// --- Siemens Structured Format ---
DATA_BLOCK "model__HS8_IW100_"
{ S7_Optimized_Access := 'TRUE' }
VERSION :
NON_RETAIN
   VAR
      W_i : ARRAY[0..7, 0..39] OF REAL;
      W_f : ARRAY[0..7, 0..39] OF REAL;
      W_g : ARRAY[0..7, 0..39] OF REAL;
      W_o : ARRAY[0..7, 0..39] OF REAL;
      R_i : ARRAY[0..7, 0..7] OF REAL;
      R_f : ARRAY[0..7, 0..7] OF REAL;
      R_g : ARRAY[0..7, 0..7] OF REAL;
      R_o : ARRAY[0..7, 0..7] OF REAL;
      B_i : ARRAY[0..7] OF REAL;
      B_f : ARRAY[0..7] OF REAL;
      B_g : ARRAY[0..7] OF REAL;
      B_o : ARRAY[0..7] OF REAL;
      FC_W : ARRAY[0..39, 0..7] OF REAL;
      FC_B : ARRAY[0..39] OF REAL;
   END_VAR
BEGIN

      W_i[0,0] := -0.00829199;
      W_i[0,1] := 0.04314763;
      W_i[0,2] := -0.00093121;
      W_i[0,3] := -0.41203406;
      W_i[0,4] := 0.14360030;
      W_i[0,5] := -0.00333697;
      W_i[0,6] := -0.05594388;
      W_i[0,7] := 0.22901678;
      W_i[0,8] := 0.12452386;
      W_i[0,9] := 0.18269505;
      W_i[0,10] := -0.00489003;
      W_i[0,11] := -1.12929618;
      W_i[0,12] := 0.50561267;
      W_i[0,13] := -0.01176495;
      W_i[0,14] := 0.05196610;
      W_i[0,15] := 0.29604533;
      W_i[0,16] := 0.00854590;
      W_i[0,17] := 0.00023653;
      W_i[0,18] := -0.05930486;
      W_i[0,19] := 0.34416831;
      W_i[0,20] := 0.04249638;
      W_i[0,21] := 0.29057521;
      W_i[0,22] := 0.00544647;
      W_i[0,23] := -0.19255431;
      W_i[0,24] := -0.20954449;
      W_i[0,25] := -0.09120649;
      W_i[0,26] := -0.00158587;
      W_i[0,27] := -0.21091045;
      W_i[0,28] := -0.00354010;
      W_i[0,29] := -0.11485449;
      W_i[0,30] := 0.40112287;
      W_i[0,31] := -0.23464951;
      W_i[0,32] := 0.07507721;
      W_i[0,33] := -0.04070815;
      W_i[0,34] := 0.16331266;
      W_i[0,35] := -0.06922071;
      W_i[0,36] := 0.07785974;
      W_i[0,37] := -0.12469714;
      W_i[0,38] := -0.09480914;
      W_i[0,39] := -0.12007505;
      W_i[1,0] := -0.14511052;
      W_i[1,1] := 0.01258339;
      W_i[1,2] := -0.02499544;
      W_i[1,3] := -0.02792050;
      W_i[1,4] := 0.05153107;
      W_i[1,5] := 0.02871069;
      W_i[1,6] := -0.00801326;
      W_i[1,7] := 0.16971111;
      W_i[1,8] := 0.07463019;
      W_i[1,9] := -0.30484986;
      W_i[1,10] := 0.00891454;
      W_i[1,11] := 0.19871780;
      W_i[1,12] := 0.02821600;
      W_i[1,13] := -0.07369927;
      W_i[1,14] := 0.02203551;
      W_i[1,15] := 0.08398883;
      W_i[1,16] := 0.00458911;
      W_i[1,17] := 0.01521466;
      W_i[1,18] := 0.06061148;
      W_i[1,19] := -0.08532640;
      W_i[1,20] := 0.01589951;
      W_i[1,21] := 0.00234504;
      W_i[1,22] := -0.04496472;
      W_i[1,23] := -0.04576229;
      W_i[1,24] := 0.03349697;
      W_i[1,25] := -0.14834076;
      W_i[1,26] := -0.00671506;
      W_i[1,27] := -0.04002256;
      W_i[1,28] := -0.05524301;
      W_i[1,29] := -0.04596998;
      W_i[1,30] := 0.20154108;
      W_i[1,31] := -0.04227936;
      W_i[1,32] := 0.27783859;
      W_i[1,33] := -0.15889524;
      W_i[1,34] := -0.17870863;
      W_i[1,35] := -0.22829576;
      W_i[1,36] := 0.00769149;
      W_i[1,37] := 0.21033208;
      W_i[1,38] := 0.02056267;
      W_i[1,39] := 0.03890164;
      W_i[2,0] := -0.00940658;
      W_i[2,1] := 0.01171005;
      W_i[2,2] := 0.01976776;
      W_i[2,3] := -0.01506334;
      W_i[2,4] := -0.01478560;
      W_i[2,5] := 0.02109193;
      W_i[2,6] := 0.01444429;
      W_i[2,7] := 0.00977760;
      W_i[2,8] := 0.06673528;
      W_i[2,9] := 0.07852798;
      W_i[2,10] := -0.02388507;
      W_i[2,11] := 0.15636960;
      W_i[2,12] := 0.04547270;
      W_i[2,13] := 0.05332979;
      W_i[2,14] := 0.02128568;
      W_i[2,15] := -0.06670643;
      W_i[2,16] := -0.00303149;
      W_i[2,17] := -0.01812665;
      W_i[2,18] := 0.09366660;
      W_i[2,19] := -0.02572775;
      W_i[2,20] := -0.02855127;
      W_i[2,21] := -0.05881069;
      W_i[2,22] := -0.05029222;
      W_i[2,23] := 0.09357284;
      W_i[2,24] := -0.46770903;
      W_i[2,25] := -0.71739095;
      W_i[2,26] := -0.03358178;
      W_i[2,27] := -0.11196791;
      W_i[2,28] := 0.12867627;
      W_i[2,29] := -0.15594745;
      W_i[2,30] := -0.02176742;
      W_i[2,31] := 0.05814255;
      W_i[2,32] := 0.02967955;
      W_i[2,33] := -0.32135192;
      W_i[2,34] := -0.70631939;
      W_i[2,35] := 0.13404904;
      W_i[2,36] := -0.05614626;
      W_i[2,37] := -0.06990065;
      W_i[2,38] := 0.09054608;
      W_i[2,39] := 0.08889610;
      W_i[3,0] := 0.05596327;
      W_i[3,1] := -0.32603350;
      W_i[3,2] := -0.13964993;
      W_i[3,3] := -0.15204740;
      W_i[3,4] := 0.05851153;
      W_i[3,5] := 0.08759125;
      W_i[3,6] := 0.07076695;
      W_i[3,7] := 0.05082684;
      W_i[3,8] := 0.00611771;
      W_i[3,9] := -0.05680722;
      W_i[3,10] := 0.04656018;
      W_i[3,11] := 0.08742622;
      W_i[3,12] := -0.00764282;
      W_i[3,13] := -0.35034382;
      W_i[3,14] := -0.12616983;
      W_i[3,15] := 0.03790347;
      W_i[3,16] := -0.00427554;
      W_i[3,17] := 0.10194600;
      W_i[3,18] := -0.06467836;
      W_i[3,19] := -0.04557304;
      W_i[3,20] := 0.13014187;
      W_i[3,21] := -0.11706656;
      W_i[3,22] := 0.20328589;
      W_i[3,23] := 0.31214345;
      W_i[3,24] := -0.19055620;
      W_i[3,25] := 0.11225392;
      W_i[3,26] := -0.00316885;
      W_i[3,27] := 0.02801218;
      W_i[3,28] := 0.07838947;
      W_i[3,29] := -0.08224142;
      W_i[3,30] := 0.02575504;
      W_i[3,31] := 0.07745822;
      W_i[3,32] := 0.05140261;
      W_i[3,33] := 0.00126193;
      W_i[3,34] := 0.03769523;
      W_i[3,35] := -0.21655150;
      W_i[3,36] := -0.08745287;
      W_i[3,37] := 0.10195030;
      W_i[3,38] := -0.44626316;
      W_i[3,39] := -0.86872011;
      W_i[4,0] := -0.04617658;
      W_i[4,1] := -0.03314103;
      W_i[4,2] := -0.08659177;
      W_i[4,3] := -0.10351395;
      W_i[4,4] := 0.06772576;
      W_i[4,5] := -0.04269263;
      W_i[4,6] := -0.04438864;
      W_i[4,7] := -0.01167864;
      W_i[4,8] := 0.02057231;
      W_i[4,9] := -0.07837452;
      W_i[4,10] := -0.03820154;
      W_i[4,11] := -0.03692231;
      W_i[4,12] := -0.07637376;
      W_i[4,13] := -0.06241865;
      W_i[4,14] := -0.01509702;
      W_i[4,15] := 0.07582836;
      W_i[4,16] := -0.01766248;
      W_i[4,17] := 0.00024068;
      W_i[4,18] := 0.03632537;
      W_i[4,19] := 0.01485146;
      W_i[4,20] := 0.10803255;
      W_i[4,21] := -0.14425407;
      W_i[4,22] := -0.01218021;
      W_i[4,23] := -0.01190184;
      W_i[4,24] := -0.46979687;
      W_i[4,25] := -0.46851084;
      W_i[4,26] := -0.02849982;
      W_i[4,27] := 0.03427306;
      W_i[4,28] := 0.04523883;
      W_i[4,29] := 0.25723371;
      W_i[4,30] := -0.09724599;
      W_i[4,31] := 0.03623974;
      W_i[4,32] := -0.10095317;
      W_i[4,33] := 0.12443283;
      W_i[4,34] := -0.42049277;
      W_i[4,35] := -0.03480925;
      W_i[4,36] := 0.04771702;
      W_i[4,37] := 0.04326405;
      W_i[4,38] := 0.03356932;
      W_i[4,39] := 0.03849664;
      W_i[5,0] := -0.17091992;
      W_i[5,1] := -0.04787771;
      W_i[5,2] := -0.02202379;
      W_i[5,3] := -0.09034166;
      W_i[5,4] := -0.00740036;
      W_i[5,5] := 0.00184778;
      W_i[5,6] := 0.01398086;
      W_i[5,7] := -0.08714975;
      W_i[5,8] := -0.10723638;
      W_i[5,9] := 0.27444202;
      W_i[5,10] := 0.02795951;
      W_i[5,11] := 0.16468486;
      W_i[5,12] := -0.25734791;
      W_i[5,13] := -0.08599530;
      W_i[5,14] := -0.07228005;
      W_i[5,15] := 0.24830806;
      W_i[5,16] := 0.04241711;
      W_i[5,17] := -0.00679267;
      W_i[5,18] := 1.35323977;
      W_i[5,19] := 0.07199069;
      W_i[5,20] := 0.06845883;
      W_i[5,21] := 0.20864677;
      W_i[5,22] := -0.14911477;
      W_i[5,23] := 0.14023533;
      W_i[5,24] := -0.02367306;
      W_i[5,25] := 0.60291624;
      W_i[5,26] := -0.19428003;
      W_i[5,27] := -0.32415670;
      W_i[5,28] := 0.17960674;
      W_i[5,29] := 0.09058087;
      W_i[5,30] := -0.24361624;
      W_i[5,31] := -0.07183243;
      W_i[5,32] := 0.01278071;
      W_i[5,33] := -0.11311200;
      W_i[5,34] := 0.64622027;
      W_i[5,35] := -0.06918935;
      W_i[5,36] := 0.04555825;
      W_i[5,37] := -0.41487035;
      W_i[5,38] := -0.02093678;
      W_i[5,39] := 0.11062510;
      W_i[6,0] := -0.08444463;
      W_i[6,1] := 0.03796263;
      W_i[6,2] := 0.02793699;
      W_i[6,3] := 0.08258326;
      W_i[6,4] := 0.01806726;
      W_i[6,5] := 0.04154406;
      W_i[6,6] := 0.06518649;
      W_i[6,7] := -0.35571000;
      W_i[6,8] := -0.08575057;
      W_i[6,9] := 0.03024576;
      W_i[6,10] := 0.08267769;
      W_i[6,11] := -0.51406556;
      W_i[6,12] := -0.18283555;
      W_i[6,13] := 0.08692829;
      W_i[6,14] := -0.01571506;
      W_i[6,15] := 0.41990465;
      W_i[6,16] := 0.06421173;
      W_i[6,17] := 0.02368255;
      W_i[6,18] := 0.00736057;
      W_i[6,19] := 0.13490863;
      W_i[6,20] := 0.24439722;
      W_i[6,21] := 0.22145407;
      W_i[6,22] := 0.23587099;
      W_i[6,23] := -0.08479463;
      W_i[6,24] := 0.15434107;
      W_i[6,25] := 0.35517022;
      W_i[6,26] := 0.02139992;
      W_i[6,27] := -0.18648548;
      W_i[6,28] := 0.00971483;
      W_i[6,29] := -0.15883411;
      W_i[6,30] := 0.16745885;
      W_i[6,31] := -0.09647866;
      W_i[6,32] := 0.20241226;
      W_i[6,33] := -0.10213183;
      W_i[6,34] := 0.35625863;
      W_i[6,35] := -0.21271712;
      W_i[6,36] := 0.07117779;
      W_i[6,37] := -0.05264070;
      W_i[6,38] := -0.07197802;
      W_i[6,39] := 0.05570221;
      W_i[7,0] := -0.14402835;
      W_i[7,1] := -0.07068059;
      W_i[7,2] := 0.04391022;
      W_i[7,3] := -0.23145308;
      W_i[7,4] := 0.01739045;
      W_i[7,5] := -0.09847571;
      W_i[7,6] := -0.07244503;
      W_i[7,7] := 0.54241705;
      W_i[7,8] := 0.05786600;
      W_i[7,9] := -0.11313851;
      W_i[7,10] := 0.05011918;
      W_i[7,11] := -0.88967866;
      W_i[7,12] := -0.78758240;
      W_i[7,13] := -0.07027908;
      W_i[7,14] := -0.15626858;
      W_i[7,15] := -0.01163841;
      W_i[7,16] := 0.06607775;
      W_i[7,17] := -0.20021817;
      W_i[7,18] := 0.08560139;
      W_i[7,19] := -0.06735905;
      W_i[7,20] := 0.11073713;
      W_i[7,21] := 0.03392316;
      W_i[7,22] := -0.07517586;
      W_i[7,23] := -0.07473031;
      W_i[7,24] := 0.17482267;
      W_i[7,25] := 0.75477821;
      W_i[7,26] := -0.19560531;
      W_i[7,27] := -0.00529976;
      W_i[7,28] := 0.06779508;
      W_i[7,29] := -0.05984003;
      W_i[7,30] := 0.36871162;
      W_i[7,31] := 0.09751310;
      W_i[7,32] := -0.32882604;
      W_i[7,33] := 0.10271895;
      W_i[7,34] := 0.03595359;
      W_i[7,35] := -0.06912012;
      W_i[7,36] := 0.05955562;
      W_i[7,37] := 0.15649518;
      W_i[7,38] := -0.16574396;
      W_i[7,39] := 0.02650662;
      W_f[0,0] := -0.08104721;
      W_f[0,1] := 0.02299085;
      W_f[0,2] := -0.08156814;
      W_f[0,3] := 0.34981409;
      W_f[0,4] := -0.02991411;
      W_f[0,5] := 0.05847026;
      W_f[0,6] := 0.08058469;
      W_f[0,7] := 0.08683547;
      W_f[0,8] := 0.02113942;
      W_f[0,9] := -0.22806560;
      W_f[0,10] := -0.04616724;
      W_f[0,11] := -0.04299140;
      W_f[0,12] := 0.11675275;
      W_f[0,13] := -0.09660369;
      W_f[0,14] := -0.04888760;
      W_f[0,15] := -0.18213840;
      W_f[0,16] := 0.12695764;
      W_f[0,17] := 0.22833031;
      W_f[0,18] := -0.03068344;
      W_f[0,19] := -0.22004378;
      W_f[0,20] := 0.01699636;
      W_f[0,21] := 0.10058182;
      W_f[0,22] := 0.02436358;
      W_f[0,23] := 0.01155086;
      W_f[0,24] := 0.67554194;
      W_f[0,25] := 0.77170414;
      W_f[0,26] := 0.04872859;
      W_f[0,27] := 0.04316394;
      W_f[0,28] := 0.01004832;
      W_f[0,29] := 0.10533538;
      W_f[0,30] := 0.26388049;
      W_f[0,31] := 0.16926253;
      W_f[0,32] := 0.31521299;
      W_f[0,33] := 0.23292090;
      W_f[0,34] := 0.71050066;
      W_f[0,35] := 0.07673426;
      W_f[0,36] := -0.03209021;
      W_f[0,37] := -0.07602870;
      W_f[0,38] := 0.07363247;
      W_f[0,39] := 0.09119339;
      W_f[1,0] := -0.02197713;
      W_f[1,1] := -0.01616614;
      W_f[1,2] := -0.02013298;
      W_f[1,3] := -0.00875140;
      W_f[1,4] := 0.04112979;
      W_f[1,5] := 0.05162001;
      W_f[1,6] := 0.00973919;
      W_f[1,7] := 0.07910040;
      W_f[1,8] := -0.31076026;
      W_f[1,9] := 0.18630370;
      W_f[1,10] := -0.00576194;
      W_f[1,11] := 0.04994554;
      W_f[1,12] := 0.05406393;
      W_f[1,13] := 0.05481998;
      W_f[1,14] := 0.01417492;
      W_f[1,15] := -0.11486354;
      W_f[1,16] := 0.22028089;
      W_f[1,17] := 0.03549247;
      W_f[1,18] := 0.07496776;
      W_f[1,19] := -0.31716284;
      W_f[1,20] := 0.02977121;
      W_f[1,21] := -0.10077871;
      W_f[1,22] := 0.29007021;
      W_f[1,23] := 0.02756922;
      W_f[1,24] := 1.14809716;
      W_f[1,25] := 1.46478581;
      W_f[1,26] := -0.01241822;
      W_f[1,27] := 0.09172244;
      W_f[1,28] := 0.01175412;
      W_f[1,29] := -0.10488217;
      W_f[1,30] := 0.00364918;
      W_f[1,31] := -0.03901139;
      W_f[1,32] := -0.08511472;
      W_f[1,33] := 0.08891900;
      W_f[1,34] := 1.39858294;
      W_f[1,35] := -0.42813861;
      W_f[1,36] := -0.00882304;
      W_f[1,37] := -0.05784527;
      W_f[1,38] := -0.13634762;
      W_f[1,39] := 0.17077002;
      W_f[2,0] := 0.01542370;
      W_f[2,1] := 0.01987428;
      W_f[2,2] := 0.00323933;
      W_f[2,3] := -0.01730455;
      W_f[2,4] := 0.06355638;
      W_f[2,5] := 0.03613569;
      W_f[2,6] := -0.01693674;
      W_f[2,7] := -0.01970888;
      W_f[2,8] := -0.06606199;
      W_f[2,9] := -0.07453630;
      W_f[2,10] := -0.00336948;
      W_f[2,11] := -0.20352897;
      W_f[2,12] := -0.10294267;
      W_f[2,13] := 0.02081121;
      W_f[2,14] := 0.06329557;
      W_f[2,15] := 0.02846926;
      W_f[2,16] := 0.06616816;
      W_f[2,17] := 0.00726432;
      W_f[2,18] := 0.04505518;
      W_f[2,19] := 0.02842713;
      W_f[2,20] := -0.00391449;
      W_f[2,21] := -0.00121696;
      W_f[2,22] := -0.17400308;
      W_f[2,23] := 0.02276708;
      W_f[2,24] := 0.26592869;
      W_f[2,25] := 0.03894256;
      W_f[2,26] := 0.12431550;
      W_f[2,27] := -0.02150069;
      W_f[2,28] := -0.05582710;
      W_f[2,29] := 0.25016540;
      W_f[2,30] := 0.01012970;
      W_f[2,31] := -0.01360032;
      W_f[2,32] := -0.07151139;
      W_f[2,33] := 0.20726912;
      W_f[2,34] := -0.33328736;
      W_f[2,35] := 0.15157171;
      W_f[2,36] := 0.01685908;
      W_f[2,37] := -0.12045209;
      W_f[2,38] := 0.01227041;
      W_f[2,39] := 0.06517339;
      W_f[3,0] := 0.47573653;
      W_f[3,1] := 0.13755870;
      W_f[3,2] := -0.08410271;
      W_f[3,3] := -0.16147336;
      W_f[3,4] := 0.10956663;
      W_f[3,5] := -0.05382008;
      W_f[3,6] := -0.09864125;
      W_f[3,7] := 0.37438312;
      W_f[3,8] := -0.31137553;
      W_f[3,9] := 0.11690006;
      W_f[3,10] := -0.16711678;
      W_f[3,11] := -0.35226113;
      W_f[3,12] := 0.14284903;
      W_f[3,13] := 0.22532572;
      W_f[3,14] := 0.31750289;
      W_f[3,15] := -0.04833202;
      W_f[3,16] := 0.04104101;
      W_f[3,17] := -0.29455543;
      W_f[3,18] := -2.66076255;
      W_f[3,19] := -0.09576055;
      W_f[3,20] := -0.16356435;
      W_f[3,21] := 0.10903085;
      W_f[3,22] := -0.44664004;
      W_f[3,23] := -0.17856193;
      W_f[3,24] := 0.41079015;
      W_f[3,25] := 0.15273106;
      W_f[3,26] := -0.33044237;
      W_f[3,27] := -0.18228154;
      W_f[3,28] := 0.04568926;
      W_f[3,29] := 1.02778792;
      W_f[3,30] := -0.34178400;
      W_f[3,31] := -0.00056406;
      W_f[3,32] := 0.21154980;
      W_f[3,33] := -0.10385001;
      W_f[3,34] := 0.03440418;
      W_f[3,35] := 0.25746328;
      W_f[3,36] := 0.02392143;
      W_f[3,37] := -0.14384723;
      W_f[3,38] := 0.40537423;
      W_f[3,39] := -0.08356514;
      W_f[4,0] := 0.01179661;
      W_f[4,1] := 0.06130485;
      W_f[4,2] := 0.00775665;
      W_f[4,3] := -0.01987305;
      W_f[4,4] := 0.03156713;
      W_f[4,5] := -0.03151586;
      W_f[4,6] := -0.06941684;
      W_f[4,7] := -0.05865467;
      W_f[4,8] := -0.12223195;
      W_f[4,9] := 0.00069460;
      W_f[4,10] := -0.01235222;
      W_f[4,11] := -0.05694751;
      W_f[4,12] := -0.00690056;
      W_f[4,13] := 0.02081548;
      W_f[4,14] := -0.02345082;
      W_f[4,15] := -0.08427138;
      W_f[4,16] := 0.00219320;
      W_f[4,17] := -0.00790089;
      W_f[4,18] := 0.06579314;
      W_f[4,19] := -0.04613130;
      W_f[4,20] := 0.06156648;
      W_f[4,21] := 0.08230194;
      W_f[4,22] := 0.02192603;
      W_f[4,23] := -0.05004644;
      W_f[4,24] := -0.33776584;
      W_f[4,25] := -0.57119745;
      W_f[4,26] := 0.00284863;
      W_f[4,27] := -0.03237003;
      W_f[4,28] := -0.06698364;
      W_f[4,29] := -0.32339925;
      W_f[4,30] := 0.06599762;
      W_f[4,31] := 0.03372506;
      W_f[4,32] := 0.20183899;
      W_f[4,33] := 0.09781818;
      W_f[4,34] := 0.21647416;
      W_f[4,35] := -0.03968338;
      W_f[4,36] := 0.04764435;
      W_f[4,37] := -0.09999206;
      W_f[4,38] := -0.04979988;
      W_f[4,39] := 0.04298165;
      W_f[5,0] := -0.00328023;
      W_f[5,1] := 0.05526555;
      W_f[5,2] := -0.02378737;
      W_f[5,3] := 0.07470135;
      W_f[5,4] := 0.07415909;
      W_f[5,5] := 0.03875844;
      W_f[5,6] := 0.04064441;
      W_f[5,7] := 0.01137258;
      W_f[5,8] := 0.04157886;
      W_f[5,9] := -0.11250745;
      W_f[5,10] := -0.03683221;
      W_f[5,11] := -0.05140235;
      W_f[5,12] := 0.16510846;
      W_f[5,13] := -0.00409127;
      W_f[5,14] := -0.03037189;
      W_f[5,15] := -0.14330336;
      W_f[5,16] := -0.02087791;
      W_f[5,17] := 0.05005715;
      W_f[5,18] := -0.06411071;
      W_f[5,19] := -0.05833034;
      W_f[5,20] := 0.00247585;
      W_f[5,21] := 0.07365038;
      W_f[5,22] := 0.00771155;
      W_f[5,23] := -0.07253324;
      W_f[5,24] := 0.94747639;
      W_f[5,25] := 0.65536422;
      W_f[5,26] := 0.01926010;
      W_f[5,27] := -0.07741715;
      W_f[5,28] := -0.02838454;
      W_f[5,29] := -0.25596547;
      W_f[5,30] := 0.04823640;
      W_f[5,31] := 0.03441899;
      W_f[5,32] := -0.04197009;
      W_f[5,33] := 0.14078745;
      W_f[5,34] := 0.25478148;
      W_f[5,35] := -0.08758619;
      W_f[5,36] := -0.00409188;
      W_f[5,37] := 0.10015804;
      W_f[5,38] := -0.01840312;
      W_f[5,39] := 0.04281899;
      W_f[6,0] := -0.03747290;
      W_f[6,1] := 0.00117479;
      W_f[6,2] := 0.01929842;
      W_f[6,3] := -0.16080324;
      W_f[6,4] := -0.00967213;
      W_f[6,5] := 0.02158868;
      W_f[6,6] := -0.07005120;
      W_f[6,7] := 0.21899310;
      W_f[6,8] := 0.03782399;
      W_f[6,9] := -0.21971041;
      W_f[6,10] := -0.04937140;
      W_f[6,11] := 0.04276552;
      W_f[6,12] := 0.02347153;
      W_f[6,13] := -0.08741955;
      W_f[6,14] := 0.02819359;
      W_f[6,15] := -0.32513508;
      W_f[6,16] := 0.09819235;
      W_f[6,17] := -0.00175993;
      W_f[6,18] := 0.00046430;
      W_f[6,19] := 0.00414359;
      W_f[6,20] := 0.05726501;
      W_f[6,21] := 0.02174316;
      W_f[6,22] := 0.40702432;
      W_f[6,23] := 0.05224282;
      W_f[6,24] := 1.36585915;
      W_f[6,25] := 1.40137434;
      W_f[6,26] := 0.06176697;
      W_f[6,27] := 0.03423437;
      W_f[6,28] := 0.01783603;
      W_f[6,29] := -0.56917655;
      W_f[6,30] := 0.47907564;
      W_f[6,31] := 0.10644426;
      W_f[6,32] := 0.44268256;
      W_f[6,33] := 0.56317347;
      W_f[6,34] := 1.12857997;
      W_f[6,35] := 0.00323946;
      W_f[6,36] := -0.03574727;
      W_f[6,37] := -0.12019916;
      W_f[6,38] := -0.04353496;
      W_f[6,39] := 0.18841393;
      W_f[7,0] := 0.08367904;
      W_f[7,1] := -0.02769166;
      W_f[7,2] := 0.05256313;
      W_f[7,3] := -0.02467708;
      W_f[7,4] := -0.08298105;
      W_f[7,5] := -0.01648388;
      W_f[7,6] := -0.04057755;
      W_f[7,7] := 0.05192674;
      W_f[7,8] := -0.03598220;
      W_f[7,9] := -0.13019682;
      W_f[7,10] := 0.01959694;
      W_f[7,11] := 0.00413586;
      W_f[7,12] := 0.05873092;
      W_f[7,13] := 0.02881050;
      W_f[7,14] := -0.02888235;
      W_f[7,15] := -0.13839944;
      W_f[7,16] := 0.02485734;
      W_f[7,17] := -0.11965133;
      W_f[7,18] := -0.11112632;
      W_f[7,19] := 0.03353542;
      W_f[7,20] := 0.02333037;
      W_f[7,21] := 0.04703392;
      W_f[7,22] := 0.20441540;
      W_f[7,23] := 0.07088239;
      W_f[7,24] := 0.59273797;
      W_f[7,25] := 0.38002837;
      W_f[7,26] := 0.01679641;
      W_f[7,27] := 0.03724186;
      W_f[7,28] := -0.06413292;
      W_f[7,29] := -0.13961390;
      W_f[7,30] := 0.11306310;
      W_f[7,31] := -0.00102062;
      W_f[7,32] := 0.19089061;
      W_f[7,33] := 0.12474129;
      W_f[7,34] := 0.52092993;
      W_f[7,35] := 0.02751438;
      W_f[7,36] := 0.01992416;
      W_f[7,37] := -0.08247742;
      W_f[7,38] := -0.05664129;
      W_f[7,39] := 0.16597328;
      W_g[0,0] := -0.06630491;
      W_g[0,1] := 0.02753393;
      W_g[0,2] := -0.06609154;
      W_g[0,3] := 0.03565337;
      W_g[0,4] := -0.14254735;
      W_g[0,5] := 0.07333323;
      W_g[0,6] := 0.14428975;
      W_g[0,7] := 0.03311217;
      W_g[0,8] := 0.02892466;
      W_g[0,9] := 0.04255950;
      W_g[0,10] := -0.03547552;
      W_g[0,11] := 0.02729788;
      W_g[0,12] := 0.02407304;
      W_g[0,13] := -0.01838484;
      W_g[0,14] := -0.04254790;
      W_g[0,15] := 0.00052823;
      W_g[0,16] := 0.02627059;
      W_g[0,17] := 0.12881427;
      W_g[0,18] := -0.04993503;
      W_g[0,19] := 0.05080932;
      W_g[0,20] := -0.13986340;
      W_g[0,21] := 0.11638415;
      W_g[0,22] := 0.01129120;
      W_g[0,23] := -0.00916141;
      W_g[0,24] := 0.20254859;
      W_g[0,25] := 0.08704451;
      W_g[0,26] := -0.03924693;
      W_g[0,27] := 0.10738914;
      W_g[0,28] := -0.04623365;
      W_g[0,29] := -0.00351558;
      W_g[0,30] := 0.00354978;
      W_g[0,31] := 0.00794905;
      W_g[0,32] := 0.00442744;
      W_g[0,33] := 0.00612418;
      W_g[0,34] := -0.20538065;
      W_g[0,35] := 0.03906323;
      W_g[0,36] := -0.00062364;
      W_g[0,37] := 0.00209236;
      W_g[0,38] := -0.03761620;
      W_g[0,39] := -0.04062740;
      W_g[1,0] := -0.10235135;
      W_g[1,1] := 0.06025442;
      W_g[1,2] := -0.09398326;
      W_g[1,3] := 0.05591756;
      W_g[1,4] := -0.10170189;
      W_g[1,5] := 0.04167721;
      W_g[1,6] := 0.01649847;
      W_g[1,7] := 0.04434075;
      W_g[1,8] := 0.04717555;
      W_g[1,9] := 0.03831566;
      W_g[1,10] := 0.05404275;
      W_g[1,11] := 0.16338016;
      W_g[1,12] := 0.15951122;
      W_g[1,13] := 0.02527176;
      W_g[1,14] := -0.01270708;
      W_g[1,15] := 0.16955729;
      W_g[1,16] := -0.08400796;
      W_g[1,17] := -0.09564576;
      W_g[1,18] := -0.16610350;
      W_g[1,19] := 0.18888752;
      W_g[1,20] := -0.02569673;
      W_g[1,21] := -0.05631816;
      W_g[1,22] := -0.01589629;
      W_g[1,23] := 0.06837284;
      W_g[1,24] := 0.19006948;
      W_g[1,25] := -0.18527375;
      W_g[1,26] := 0.06264018;
      W_g[1,27] := -0.06131431;
      W_g[1,28] := -0.02992554;
      W_g[1,29] := 0.02249875;
      W_g[1,30] := -0.01341370;
      W_g[1,31] := -0.01471063;
      W_g[1,32] := -0.01641031;
      W_g[1,33] := -0.02138708;
      W_g[1,34] := 0.09338091;
      W_g[1,35] := 0.17898178;
      W_g[1,36] := -0.08693415;
      W_g[1,37] := -0.19239108;
      W_g[1,38] := -0.05011347;
      W_g[1,39] := -0.03428216;
      W_g[2,0] := 0.06590919;
      W_g[2,1] := 0.01555668;
      W_g[2,2] := 0.05944061;
      W_g[2,3] := -0.00003379;
      W_g[2,4] := -0.16144016;
      W_g[2,5] := 0.07584924;
      W_g[2,6] := 0.07926709;
      W_g[2,7] := 0.00562621;
      W_g[2,8] := 0.00176247;
      W_g[2,9] := 0.00667630;
      W_g[2,10] := -0.01289325;
      W_g[2,11] := -0.03508691;
      W_g[2,12] := -0.03598065;
      W_g[2,13] := 0.14380608;
      W_g[2,14] := 0.06675316;
      W_g[2,15] := -0.02170967;
      W_g[2,16] := 0.03013330;
      W_g[2,17] := -0.04029799;
      W_g[2,18] := -0.14855465;
      W_g[2,19] := 0.00260400;
      W_g[2,20] := -0.08315958;
      W_g[2,21] := 0.01309617;
      W_g[2,22] := 0.05792306;
      W_g[2,23] := 0.14916992;
      W_g[2,24] := 0.13496941;
      W_g[2,25] := 0.20256528;
      W_g[2,26] := 0.06222376;
      W_g[2,27] := 0.00734210;
      W_g[2,28] := -0.04847896;
      W_g[2,29] := -0.00581570;
      W_g[2,30] := 0.03206468;
      W_g[2,31] := 0.02264830;
      W_g[2,32] := 0.04472146;
      W_g[2,33] := 0.04833479;
      W_g[2,34] := 0.68682790;
      W_g[2,35] := 0.03641244;
      W_g[2,36] := -0.05233013;
      W_g[2,37] := 0.01984018;
      W_g[2,38] := 0.05872162;
      W_g[2,39] := 0.05237507;
      W_g[3,0] := -0.05719843;
      W_g[3,1] := 0.06765803;
      W_g[3,2] := -0.05017579;
      W_g[3,3] := -0.09871275;
      W_g[3,4] := -0.14791933;
      W_g[3,5] := -0.05363221;
      W_g[3,6] := -0.11064304;
      W_g[3,7] := -0.06622731;
      W_g[3,8] := -0.06549069;
      W_g[3,9] := -0.07995880;
      W_g[3,10] := -0.00412930;
      W_g[3,11] := -0.05527864;
      W_g[3,12] := -0.05236278;
      W_g[3,13] := 0.01281861;
      W_g[3,14] := 0.00663725;
      W_g[3,15] := -0.05022956;
      W_g[3,16] := 0.00247445;
      W_g[3,17] := -0.00537014;
      W_g[3,18] := -0.17336990;
      W_g[3,19] := -0.04672612;
      W_g[3,20] := 0.08145336;
      W_g[3,21] := 0.04289828;
      W_g[3,22] := -0.04270948;
      W_g[3,23] := -0.00124830;
      W_g[3,24] := -0.58283401;
      W_g[3,25] := -0.74716926;
      W_g[3,26] := -0.05420419;
      W_g[3,27] := 0.04391639;
      W_g[3,28] := -0.21304598;
      W_g[3,29] := 0.14126062;
      W_g[3,30] := -0.04634099;
      W_g[3,31] := -0.01238058;
      W_g[3,32] := -0.02521331;
      W_g[3,33] := -0.01312026;
      W_g[3,34] := 0.00096928;
      W_g[3,35] := -0.08583874;
      W_g[3,36] := 0.04279795;
      W_g[3,37] := 0.07323888;
      W_g[3,38] := -0.00020507;
      W_g[3,39] := 0.48666921;
      W_g[4,0] := 0.03492008;
      W_g[4,1] := -0.06098935;
      W_g[4,2] := 0.03832612;
      W_g[4,3] := 0.05924186;
      W_g[4,4] := -0.04744076;
      W_g[4,5] := 0.03529921;
      W_g[4,6] := 0.07721187;
      W_g[4,7] := 0.05416005;
      W_g[4,8] := 0.05382877;
      W_g[4,9] := 0.06243544;
      W_g[4,10] := 0.00853686;
      W_g[4,11] := -0.00808500;
      W_g[4,12] := -0.00045702;
      W_g[4,13] := -0.01504347;
      W_g[4,14] := 0.05096063;
      W_g[4,15] := 0.00273409;
      W_g[4,16] := 0.04891136;
      W_g[4,17] := 0.01359798;
      W_g[4,18] := -0.04669548;
      W_g[4,19] := 0.01079443;
      W_g[4,20] := -0.08128674;
      W_g[4,21] := 0.02045462;
      W_g[4,22] := -0.03726062;
      W_g[4,23] := 0.01082981;
      W_g[4,24] := -0.72472757;
      W_g[4,25] := -0.60457122;
      W_g[4,26] := -0.02546896;
      W_g[4,27] := 0.02074758;
      W_g[4,28] := 0.02423066;
      W_g[4,29] := 0.02050022;
      W_g[4,30] := -0.03584260;
      W_g[4,31] := -0.03780675;
      W_g[4,32] := -0.01639182;
      W_g[4,33] := -0.01888406;
      W_g[4,34] := -0.90565455;
      W_g[4,35] := -0.02123658;
      W_g[4,36] := -0.05081832;
      W_g[4,37] := -0.08846542;
      W_g[4,38] := 0.05660410;
      W_g[4,39] := 0.05612533;
      W_g[5,0] := 0.11782174;
      W_g[5,1] := -0.06627837;
      W_g[5,2] := 0.11258242;
      W_g[5,3] := -0.00078306;
      W_g[5,4] := -0.06244962;
      W_g[5,5] := -0.05785579;
      W_g[5,6] := -0.07869791;
      W_g[5,7] := 0.01213171;
      W_g[5,8] := 0.00927653;
      W_g[5,9] := 0.00150932;
      W_g[5,10] := 0.04006030;
      W_g[5,11] := -0.02427769;
      W_g[5,12] := -0.03185246;
      W_g[5,13] := 0.04451595;
      W_g[5,14] := -0.07225010;
      W_g[5,15] := -0.01958377;
      W_g[5,16] := -0.07384533;
      W_g[5,17] := -0.05695982;
      W_g[5,18] := 0.01737016;
      W_g[5,19] := -0.04037121;
      W_g[5,20] := 0.06191914;
      W_g[5,21] := 0.01803040;
      W_g[5,22] := -0.01919131;
      W_g[5,23] := 0.05039211;
      W_g[5,24] := -0.12293056;
      W_g[5,25] := 0.30277607;
      W_g[5,26] := -0.03416682;
      W_g[5,27] := 0.04258297;
      W_g[5,28] := -0.09654819;
      W_g[5,29] := 0.03460327;
      W_g[5,30] := -0.02886237;
      W_g[5,31] := -0.00133085;
      W_g[5,32] := -0.02660071;
      W_g[5,33] := -0.00949432;
      W_g[5,34] := -0.00906071;
      W_g[5,35] := -0.07421639;
      W_g[5,36] := 0.04989494;
      W_g[5,37] := 0.06070245;
      W_g[5,38] := -0.07028808;
      W_g[5,39] := -0.06729650;
      W_g[6,0] := 0.05034672;
      W_g[6,1] := 0.00489272;
      W_g[6,2] := 0.04725259;
      W_g[6,3] := -0.08067816;
      W_g[6,4] := 0.00670493;
      W_g[6,5] := 0.08702958;
      W_g[6,6] := 0.11027312;
      W_g[6,7] := -0.09004638;
      W_g[6,8] := -0.08810285;
      W_g[6,9] := -0.08126769;
      W_g[6,10] := -0.12583737;
      W_g[6,11] := -0.01801138;
      W_g[6,12] := -0.02720401;
      W_g[6,13] := 0.03163574;
      W_g[6,14] := -0.01812004;
      W_g[6,15] := 0.00238652;
      W_g[6,16] := -0.08167886;
      W_g[6,17] := -0.11650438;
      W_g[6,18] := 0.00859512;
      W_g[6,19] := -0.03721597;
      W_g[6,20] := -0.11230972;
      W_g[6,21] := 0.03647594;
      W_g[6,22] := -0.00780440;
      W_g[6,23] := -0.02305741;
      W_g[6,24] := -0.15329531;
      W_g[6,25] := -0.10199876;
      W_g[6,26] := -0.01837613;
      W_g[6,27] := 0.03090143;
      W_g[6,28] := 0.10385493;
      W_g[6,29] := -0.01681059;
      W_g[6,30] := 0.00302486;
      W_g[6,31] := -0.01577753;
      W_g[6,32] := 0.00630172;
      W_g[6,33] := -0.00393950;
      W_g[6,34] := 0.11279012;
      W_g[6,35] := -0.00852283;
      W_g[6,36] := -0.02479460;
      W_g[6,37] := -0.03145938;
      W_g[6,38] := -0.03585445;
      W_g[6,39] := -0.02777989;
      W_g[7,0] := 0.02680640;
      W_g[7,1] := -0.00984313;
      W_g[7,2] := 0.02535466;
      W_g[7,3] := -0.00817555;
      W_g[7,4] := 0.06542997;
      W_g[7,5] := 0.00822230;
      W_g[7,6] := -0.01459355;
      W_g[7,7] := -0.01140613;
      W_g[7,8] := -0.00660438;
      W_g[7,9] := -0.00928965;
      W_g[7,10] := 0.00062967;
      W_g[7,11] := -0.07829287;
      W_g[7,12] := -0.05349097;
      W_g[7,13] := 0.02648462;
      W_g[7,14] := -0.05610063;
      W_g[7,15] := -0.07086886;
      W_g[7,16] := 0.01190711;
      W_g[7,17] := 0.09898359;
      W_g[7,18] := -0.02487384;
      W_g[7,19] := -0.05087938;
      W_g[7,20] := 0.01285185;
      W_g[7,21] := -0.06452682;
      W_g[7,22] := -0.00034817;
      W_g[7,23] := 0.01669965;
      W_g[7,24] := -0.43177298;
      W_g[7,25] := -0.03666652;
      W_g[7,26] := 0.03783032;
      W_g[7,27] := -0.06900723;
      W_g[7,28] := 0.05982220;
      W_g[7,29] := -0.03167899;
      W_g[7,30] := 0.00115681;
      W_g[7,31] := -0.00686107;
      W_g[7,32] := 0.00279485;
      W_g[7,33] := -0.00087522;
      W_g[7,34] := -0.00795635;
      W_g[7,35] := -0.00445508;
      W_g[7,36] := -0.04221371;
      W_g[7,37] := -0.02763689;
      W_g[7,38] := -0.04380527;
      W_g[7,39] := -0.04690089;
      W_o[0,0] := 0.53019369;
      W_o[0,1] := -0.06155616;
      W_o[0,2] := -0.38640434;
      W_o[0,3] := -0.15764126;
      W_o[0,4] := 0.41086245;
      W_o[0,5] := -0.03151236;
      W_o[0,6] := 0.00634237;
      W_o[0,7] := -0.13995783;
      W_o[0,8] := 0.08930115;
      W_o[0,9] := -0.02128680;
      W_o[0,10] := 0.09999584;
      W_o[0,11] := 0.10780117;
      W_o[0,12] := -0.15695846;
      W_o[0,13] := -0.18406366;
      W_o[0,14] := -0.28228819;
      W_o[0,15] := -0.51441675;
      W_o[0,16] := -0.11759740;
      W_o[0,17] := 0.32924205;
      W_o[0,18] := 1.02407587;
      W_o[0,19] := -0.14473118;
      W_o[0,20] := 0.12380417;
      W_o[0,21] := -0.00890757;
      W_o[0,22] := 0.18995185;
      W_o[0,23] := -0.02388396;
      W_o[0,24] := 1.01688302;
      W_o[0,25] := 1.32019973;
      W_o[0,26] := 0.01054627;
      W_o[0,27] := -0.38473883;
      W_o[0,28] := 0.03367974;
      W_o[0,29] := -0.04755234;
      W_o[0,30] := -0.03527200;
      W_o[0,31] := -0.08217989;
      W_o[0,32] := -0.12496393;
      W_o[0,33] := -0.15572555;
      W_o[0,34] := 1.43245482;
      W_o[0,35] := -0.10994142;
      W_o[0,36] := 0.02894684;
      W_o[0,37] := 0.02606086;
      W_o[0,38] := -0.00497870;
      W_o[0,39] := -0.02025986;
      W_o[1,0] := -0.03733223;
      W_o[1,1] := -0.05743759;
      W_o[1,2] := -0.27563941;
      W_o[1,3] := -0.02681245;
      W_o[1,4] := -0.09759782;
      W_o[1,5] := 0.03597067;
      W_o[1,6] := 0.17622416;
      W_o[1,7] := -0.28184685;
      W_o[1,8] := 0.28251758;
      W_o[1,9] := 0.40479794;
      W_o[1,10] := -0.00874605;
      W_o[1,11] := -0.22345169;
      W_o[1,12] := -0.39604142;
      W_o[1,13] := 0.13460745;
      W_o[1,14] := -0.16698690;
      W_o[1,15] := -0.29505059;
      W_o[1,16] := 0.08361635;
      W_o[1,17] := -0.35688013;
      W_o[1,18] := 0.51315767;
      W_o[1,19] := -1.03348815;
      W_o[1,20] := -0.10220779;
      W_o[1,21] := -0.18512122;
      W_o[1,22] := 0.01154257;
      W_o[1,23] := 0.09604655;
      W_o[1,24] := 1.55665982;
      W_o[1,25] := 1.30720556;
      W_o[1,26] := -0.15147182;
      W_o[1,27] := 0.07709698;
      W_o[1,28] := 0.10548013;
      W_o[1,29] := -0.07245205;
      W_o[1,30] := 0.48158705;
      W_o[1,31] := 0.21815035;
      W_o[1,32] := -0.00193443;
      W_o[1,33] := -0.17135660;
      W_o[1,34] := 0.48604634;
      W_o[1,35] := 0.38598192;
      W_o[1,36] := 0.08623584;
      W_o[1,37] := -0.08203863;
      W_o[1,38] := 0.23385969;
      W_o[1,39] := 0.42781851;
      W_o[2,0] := 0.00399225;
      W_o[2,1] := -0.05571604;
      W_o[2,2] := -0.02511727;
      W_o[2,3] := 0.02144472;
      W_o[2,4] := 0.02344707;
      W_o[2,5] := -0.08246233;
      W_o[2,6] := -0.01497909;
      W_o[2,7] := 0.02220178;
      W_o[2,8] := -0.06884211;
      W_o[2,9] := -0.09796878;
      W_o[2,10] := 0.24016623;
      W_o[2,11] := 0.10531332;
      W_o[2,12] := -0.05697370;
      W_o[2,13] := -0.11412688;
      W_o[2,14] := 0.00882436;
      W_o[2,15] := 0.01609431;
      W_o[2,16] := -0.00689903;
      W_o[2,17] := -0.02796670;
      W_o[2,18] := 1.35730100;
      W_o[2,19] := -0.02292132;
      W_o[2,20] := 0.30487630;
      W_o[2,21] := 0.05938051;
      W_o[2,22] := 0.16648391;
      W_o[2,23] := -0.45096326;
      W_o[2,24] := -0.29668695;
      W_o[2,25] := 0.11092938;
      W_o[2,26] := 0.03940877;
      W_o[2,27] := -0.05482103;
      W_o[2,28] := 0.22729106;
      W_o[2,29] := -0.04754604;
      W_o[2,30] := 0.10846881;
      W_o[2,31] := -0.04006886;
      W_o[2,32] := -0.02904707;
      W_o[2,33] := 0.33994037;
      W_o[2,34] := 0.19743054;
      W_o[2,35] := -0.01746079;
      W_o[2,36] := -0.08904223;
      W_o[2,37] := -0.22370100;
      W_o[2,38] := -0.07259841;
      W_o[2,39] := 0.63436109;
      W_o[3,0] := -0.57580048;
      W_o[3,1] := 0.07226373;
      W_o[3,2] := -0.34274739;
      W_o[3,3] := -0.13415729;
      W_o[3,4] := -0.02352028;
      W_o[3,5] := 0.01078554;
      W_o[3,6] := -0.11286568;
      W_o[3,7] := 0.00544936;
      W_o[3,8] := -0.03946435;
      W_o[3,9] := -0.23858593;
      W_o[3,10] := -0.12877348;
      W_o[3,11] := 0.23244406;
      W_o[3,12] := -0.14977308;
      W_o[3,13] := 0.15883800;
      W_o[3,14] := 0.00308700;
      W_o[3,15] := 0.02639855;
      W_o[3,16] := -0.00433945;
      W_o[3,17] := 0.02282741;
      W_o[3,18] := 0.58263451;
      W_o[3,19] := -0.00315157;
      W_o[3,20] := -0.06576378;
      W_o[3,21] := 0.25107187;
      W_o[3,22] := -0.20083913;
      W_o[3,23] := 0.15694763;
      W_o[3,24] := -0.04683150;
      W_o[3,25] := 0.02712667;
      W_o[3,26] := 0.22781134;
      W_o[3,27] := -0.33466589;
      W_o[3,28] := 0.11372802;
      W_o[3,29] := 0.13145071;
      W_o[3,30] := -0.10182201;
      W_o[3,31] := -0.22603890;
      W_o[3,32] := -0.15764055;
      W_o[3,33] := 0.47687146;
      W_o[3,34] := 0.03133727;
      W_o[3,35] := -0.15790868;
      W_o[3,36] := 0.01756845;
      W_o[3,37] := -0.13447653;
      W_o[3,38] := 0.10869049;
      W_o[3,39] := 0.03116553;
      W_o[4,0] := 0.32478511;
      W_o[4,1] := 0.26212886;
      W_o[4,2] := 0.14959159;
      W_o[4,3] := 0.00132887;
      W_o[4,4] := 0.63797754;
      W_o[4,5] := 0.56880975;
      W_o[4,6] := 0.54416990;
      W_o[4,7] := 0.04824677;
      W_o[4,8] := 0.06277762;
      W_o[4,9] := 0.34240499;
      W_o[4,10] := 0.11181158;
      W_o[4,11] := 0.25369734;
      W_o[4,12] := -0.06000311;
      W_o[4,13] := -0.15960956;
      W_o[4,14] := 0.05395936;
      W_o[4,15] := 0.00129215;
      W_o[4,16] := -0.13032414;
      W_o[4,17] := -0.05327151;
      W_o[4,18] := -0.15177877;
      W_o[4,19] := -0.25642666;
      W_o[4,20] := 0.16041021;
      W_o[4,21] := 0.17214362;
      W_o[4,22] := -0.16869369;
      W_o[4,23] := -0.02294435;
      W_o[4,24] := -0.23875684;
      W_o[4,25] := -0.16617161;
      W_o[4,26] := -0.09589908;
      W_o[4,27] := 0.08004687;
      W_o[4,28] := -0.38547710;
      W_o[4,29] := -0.13680306;
      W_o[4,30] := -0.54162902;
      W_o[4,31] := 0.18120638;
      W_o[4,32] := 0.06826349;
      W_o[4,33] := 0.20314606;
      W_o[4,34] := 0.22013944;
      W_o[4,35] := -0.04085778;
      W_o[4,36] := -0.08718784;
      W_o[4,37] := 0.08242843;
      W_o[4,38] := -0.10997366;
      W_o[4,39] := 0.13200577;
      W_o[5,0] := 0.11899070;
      W_o[5,1] := -0.37417474;
      W_o[5,2] := -0.07908265;
      W_o[5,3] := -0.20581923;
      W_o[5,4] := -0.22015102;
      W_o[5,5] := -0.01878908;
      W_o[5,6] := -0.32002872;
      W_o[5,7] := 0.03229008;
      W_o[5,8] := -0.67315555;
      W_o[5,9] := -0.18006264;
      W_o[5,10] := 0.12544481;
      W_o[5,11] := -0.29003429;
      W_o[5,12] := -0.62917036;
      W_o[5,13] := 0.04711899;
      W_o[5,14] := 0.10358876;
      W_o[5,15] := -0.37413913;
      W_o[5,16] := -0.50427359;
      W_o[5,17] := -0.04341435;
      W_o[5,18] := 0.54133219;
      W_o[5,19] := 0.16898222;
      W_o[5,20] := 0.07634972;
      W_o[5,21] := 0.15058914;
      W_o[5,22] := -0.07847997;
      W_o[5,23] := 0.12143426;
      W_o[5,24] := 1.72363305;
      W_o[5,25] := 1.55727899;
      W_o[5,26] := -0.27936074;
      W_o[5,27] := -0.02814472;
      W_o[5,28] := -0.12525134;
      W_o[5,29] := -0.13958108;
      W_o[5,30] := 0.14886966;
      W_o[5,31] := 0.02737931;
      W_o[5,32] := 0.34065816;
      W_o[5,33] := -0.18217729;
      W_o[5,34] := 0.56298286;
      W_o[5,35] := -0.12124423;
      W_o[5,36] := 0.06491477;
      W_o[5,37] := 0.01750619;
      W_o[5,38] := -0.13162488;
      W_o[5,39] := 0.77068377;
      W_o[6,0] := 0.05337723;
      W_o[6,1] := -0.10503292;
      W_o[6,2] := -0.12059452;
      W_o[6,3] := -0.07529414;
      W_o[6,4] := 0.07955431;
      W_o[6,5] := 0.14899205;
      W_o[6,6] := 1.74876642;
      W_o[6,7] := -0.00885175;
      W_o[6,8] := 0.25503284;
      W_o[6,9] := 0.02846204;
      W_o[6,10] := 0.19950083;
      W_o[6,11] := -0.32499984;
      W_o[6,12] := 0.34918392;
      W_o[6,13] := -0.10124896;
      W_o[6,14] := 0.02444035;
      W_o[6,15] := 0.01967154;
      W_o[6,16] := 0.17250372;
      W_o[6,17] := 0.12925944;
      W_o[6,18] := -0.04913221;
      W_o[6,19] := -0.12923992;
      W_o[6,20] := -0.66172892;
      W_o[6,21] := 0.14941704;
      W_o[6,22] := -0.08255627;
      W_o[6,23] := -0.17822625;
      W_o[6,24] := 1.63026547;
      W_o[6,25] := 1.15676641;
      W_o[6,26] := 0.00649359;
      W_o[6,27] := -0.09291494;
      W_o[6,28] := 0.32158482;
      W_o[6,29] := 0.00866020;
      W_o[6,30] := 0.05388094;
      W_o[6,31] := -0.07712737;
      W_o[6,32] := -0.02376380;
      W_o[6,33] := -0.14076465;
      W_o[6,34] := 1.72388208;
      W_o[6,35] := -0.06460242;
      W_o[6,36] := -0.03571915;
      W_o[6,37] := -0.00976443;
      W_o[6,38] := -0.05740520;
      W_o[6,39] := 0.81725025;
      W_o[7,0] := -0.01940660;
      W_o[7,1] := 0.01618135;
      W_o[7,2] := -0.01165283;
      W_o[7,3] := 0.10612590;
      W_o[7,4] := 0.20484668;
      W_o[7,5] := -0.04044059;
      W_o[7,6] := 0.02525332;
      W_o[7,7] := -0.03475735;
      W_o[7,8] := 0.07170975;
      W_o[7,9] := -0.01410048;
      W_o[7,10] := -0.05771373;
      W_o[7,11] := -0.41994172;
      W_o[7,12] := 0.83318508;
      W_o[7,13] := -0.10440679;
      W_o[7,14] := -0.12772350;
      W_o[7,15] := 0.10942663;
      W_o[7,16] := -0.06550087;
      W_o[7,17] := 0.33426768;
      W_o[7,18] := 0.33965129;
      W_o[7,19] := 0.45627210;
      W_o[7,20] := 0.11828049;
      W_o[7,21] := 0.40228167;
      W_o[7,22] := 0.06733994;
      W_o[7,23] := -0.22098058;
      W_o[7,24] := 1.70450640;
      W_o[7,25] := 1.64259458;
      W_o[7,26] := -0.14286987;
      W_o[7,27] := -0.55151159;
      W_o[7,28] := -0.09025964;
      W_o[7,29] := 0.02003895;
      W_o[7,30] := 0.31637633;
      W_o[7,31] := 0.08442478;
      W_o[7,32] := -0.01943155;
      W_o[7,33] := 0.12002160;
      W_o[7,34] := -0.18836913;
      W_o[7,35] := 0.32384491;
      W_o[7,36] := 0.06107497;
      W_o[7,37] := 0.26500893;
      W_o[7,38] := 0.11114403;
      W_o[7,39] := 0.78508574;
      R_i[0,0] := -1.76221621;
      R_i[0,1] := 0.52157736;
      R_i[0,2] := 0.82397699;
      R_i[0,3] := 0.23320295;
      R_i[0,4] := 0.26695707;
      R_i[0,5] := -0.39557868;
      R_i[0,6] := 0.60933948;
      R_i[0,7] := -0.90380085;
      R_i[1,0] := -0.05309208;
      R_i[1,1] := 0.13526984;
      R_i[1,2] := 0.07049563;
      R_i[1,3] := 0.22406499;
      R_i[1,4] := 1.02717400;
      R_i[1,5] := 0.37673113;
      R_i[1,6] := -0.09311269;
      R_i[1,7] := 0.54050368;
      R_i[2,0] := 0.60295075;
      R_i[2,1] := -0.28946203;
      R_i[2,2] := -1.74857521;
      R_i[2,3] := 1.08004105;
      R_i[2,4] := 0.55615216;
      R_i[2,5] := 0.56903708;
      R_i[2,6] := 0.44092867;
      R_i[2,7] := -0.19400248;
      R_i[3,0] := 0.43188563;
      R_i[3,1] := -1.42421794;
      R_i[3,2] := -0.02847767;
      R_i[3,3] := -0.64828926;
      R_i[3,4] := -0.10517685;
      R_i[3,5] := -0.59241074;
      R_i[3,6] := 0.45091745;
      R_i[3,7] := -1.67551839;
      R_i[4,0] := 0.07754488;
      R_i[4,1] := 0.48348141;
      R_i[4,2] := 0.40796608;
      R_i[4,3] := 0.50797224;
      R_i[4,4] := 0.88376588;
      R_i[4,5] := 0.46888179;
      R_i[4,6] := 0.24384692;
      R_i[4,7] := 0.24219359;
      R_i[5,0] := -0.13315447;
      R_i[5,1] := -0.18462478;
      R_i[5,2] := 0.59829623;
      R_i[5,3] := 0.34677979;
      R_i[5,4] := 0.06675477;
      R_i[5,5] := 0.68211377;
      R_i[5,6] := -0.00705162;
      R_i[5,7] := 0.06832804;
      R_i[6,0] := -0.00113238;
      R_i[6,1] := 0.62419927;
      R_i[6,2] := -0.12593758;
      R_i[6,3] := 0.19382173;
      R_i[6,4] := 1.07807183;
      R_i[6,5] := 0.30431101;
      R_i[6,6] := -0.06325435;
      R_i[6,7] := 0.48427039;
      R_i[7,0] := 0.01406168;
      R_i[7,1] := 0.75736505;
      R_i[7,2] := 1.03017557;
      R_i[7,3] := 1.73858941;
      R_i[7,4] := 0.14469253;
      R_i[7,5] := 0.04086954;
      R_i[7,6] := 0.97912145;
      R_i[7,7] := 1.66612554;
      R_f[0,0] := -0.78480172;
      R_f[0,1] := 1.04719555;
      R_f[0,2] := 0.36177492;
      R_f[0,3] := -0.28844494;
      R_f[0,4] := -1.00501108;
      R_f[0,5] := 0.86008644;
      R_f[0,6] := 0.95452124;
      R_f[0,7] := -0.42550567;
      R_f[1,0] := 0.15893026;
      R_f[1,1] := 1.37443113;
      R_f[1,2] := 0.47152451;
      R_f[1,3] := -0.38653737;
      R_f[1,4] := -1.46660495;
      R_f[1,5] := 0.14477186;
      R_f[1,6] := 0.51057285;
      R_f[1,7] := 0.11357135;
      R_f[2,0] := 0.80281532;
      R_f[2,1] := 0.70828509;
      R_f[2,2] := -0.94942558;
      R_f[2,3] := 0.11890656;
      R_f[2,4] := 0.67991215;
      R_f[2,5] := 0.77881575;
      R_f[2,6] := 0.16744818;
      R_f[2,7] := -0.15003739;
      R_f[3,0] := 1.34650016;
      R_f[3,1] := 1.08039427;
      R_f[3,2] := 0.34709018;
      R_f[3,3] := 0.39212197;
      R_f[3,4] := -0.85905784;
      R_f[3,5] := -0.47246596;
      R_f[3,6] := -0.98672587;
      R_f[3,7] := 1.46773016;
      R_f[4,0] := 0.28010875;
      R_f[4,1] := 0.40872636;
      R_f[4,2] := 0.94696331;
      R_f[4,3] := -0.99466449;
      R_f[4,4] := 0.36566308;
      R_f[4,5] := -0.05359131;
      R_f[4,6] := -0.31528312;
      R_f[4,7] := 0.03403832;
      R_f[5,0] := -0.27811784;
      R_f[5,1] := -0.04785284;
      R_f[5,2] := 0.54444504;
      R_f[5,3] := -0.26260680;
      R_f[5,4] := -0.05670305;
      R_f[5,5] := 0.03130004;
      R_f[5,6] := -0.27105442;
      R_f[5,7] := -0.42530912;
      R_f[6,0] := 0.39771050;
      R_f[6,1] := 0.86197048;
      R_f[6,2] := -0.29826346;
      R_f[6,3] := -1.11406517;
      R_f[6,4] := -0.61089790;
      R_f[6,5] := 0.83620089;
      R_f[6,6] := 0.18404177;
      R_f[6,7] := -0.26641241;
      R_f[7,0] := 0.52239841;
      R_f[7,1] := 0.12579544;
      R_f[7,2] := -0.14314617;
      R_f[7,3] := -0.70179570;
      R_f[7,4] := -0.48279399;
      R_f[7,5] := -0.67025268;
      R_f[7,6] := -0.24483326;
      R_f[7,7] := 0.38481027;
      R_g[0,0] := -2.31126142;
      R_g[0,1] := 0.15979449;
      R_g[0,2] := -0.71282071;
      R_g[0,3] := 0.53335387;
      R_g[0,4] := 0.22411184;
      R_g[0,5] := -0.22383350;
      R_g[0,6] := -0.32874081;
      R_g[0,7] := 0.17022361;
      R_g[1,0] := 0.09345370;
      R_g[1,1] := -2.93099284;
      R_g[1,2] := 0.02507862;
      R_g[1,3] := -1.16432595;
      R_g[1,4] := -0.54074705;
      R_g[1,5] := 0.00950189;
      R_g[1,6] := -0.05821744;
      R_g[1,7] := -0.14515182;
      R_g[2,0] := 0.50597680;
      R_g[2,1] := 0.14804667;
      R_g[2,2] := -3.28287935;
      R_g[2,3] := 0.89723355;
      R_g[2,4] := 0.69730288;
      R_g[2,5] := 0.14443779;
      R_g[2,6] := 0.26224744;
      R_g[2,7] := -0.06217655;
      R_g[3,0] := -0.07626731;
      R_g[3,1] := 0.18686098;
      R_g[3,2] := 0.07488978;
      R_g[3,3] := -2.59162259;
      R_g[3,4] := 0.08314367;
      R_g[3,5] := -0.03698634;
      R_g[3,6] := -0.04303954;
      R_g[3,7] := 0.13465340;
      R_g[4,0] := 0.13933653;
      R_g[4,1] := 0.01768548;
      R_g[4,2] := 0.68640625;
      R_g[4,3] := -0.88957936;
      R_g[4,4] := -3.32161546;
      R_g[4,5] := -0.09063296;
      R_g[4,6] := 0.16870818;
      R_g[4,7] := 0.07515577;
      R_g[5,0] := 0.15696557;
      R_g[5,1] := -0.32806566;
      R_g[5,2] := 0.21851663;
      R_g[5,3] := 0.00382882;
      R_g[5,4] := 0.18182336;
      R_g[5,5] := -1.54942656;
      R_g[5,6] := -0.03786261;
      R_g[5,7] := -0.40736923;
      R_g[6,0] := 0.25247186;
      R_g[6,1] := -0.21546571;
      R_g[6,2] := 0.71766186;
      R_g[6,3] := -1.00176036;
      R_g[6,4] := -0.80685157;
      R_g[6,5] := 0.03523477;
      R_g[6,6] := -2.34571934;
      R_g[6,7] := -0.16209392;
      R_g[7,0] := 0.33655006;
      R_g[7,1] := -0.20172799;
      R_g[7,2] := 0.18418945;
      R_g[7,3] := -0.82496607;
      R_g[7,4] := -0.49587831;
      R_g[7,5] := 0.11657711;
      R_g[7,6] := 0.07683489;
      R_g[7,7] := -1.71039522;
      R_o[0,0] := -0.07976321;
      R_o[0,1] := -0.28596640;
      R_o[0,2] := 0.44985750;
      R_o[0,3] := -0.04182919;
      R_o[0,4] := -0.08931469;
      R_o[0,5] := 0.22835432;
      R_o[0,6] := -0.48113039;
      R_o[0,7] := 0.45420447;
      R_o[1,0] := -0.40337405;
      R_o[1,1] := 1.10107327;
      R_o[1,2] := 0.34227836;
      R_o[1,3] := 0.63772434;
      R_o[1,4] := -1.29314208;
      R_o[1,5] := 0.62262118;
      R_o[1,6] := -0.27958676;
      R_o[1,7] := 0.91118693;
      R_o[2,0] := 0.01233310;
      R_o[2,1] := 0.40857324;
      R_o[2,2] := 3.45338154;
      R_o[2,3] := -0.72523892;
      R_o[2,4] := -0.55717379;
      R_o[2,5] := 0.02638322;
      R_o[2,6] := -0.03600628;
      R_o[2,7] := 0.75784165;
      R_o[3,0] := 0.55902964;
      R_o[3,1] := -0.39030707;
      R_o[3,2] := 1.01299071;
      R_o[3,3] := -2.74955440;
      R_o[3,4] := -1.36864233;
      R_o[3,5] := -0.26874191;
      R_o[3,6] := 0.12407675;
      R_o[3,7] := -0.44909188;
      R_o[4,0] := 0.12900312;
      R_o[4,1] := 0.75504678;
      R_o[4,2] := 2.00499749;
      R_o[4,3] := -0.11805858;
      R_o[4,4] := -2.42332268;
      R_o[4,5] := -0.78491461;
      R_o[4,6] := -0.11813148;
      R_o[4,7] := 0.26362744;
      R_o[5,0] := 0.77286434;
      R_o[5,1] := 0.76400870;
      R_o[5,2] := 0.76163286;
      R_o[5,3] := 0.25209603;
      R_o[5,4] := -0.85733461;
      R_o[5,5] := -0.87099206;
      R_o[5,6] := 0.31007352;
      R_o[5,7] := 0.03706209;
      R_o[6,0] := 0.18698657;
      R_o[6,1] := -0.21811183;
      R_o[6,2] := 1.00948119;
      R_o[6,3] := 0.17257449;
      R_o[6,4] := -0.63534433;
      R_o[6,5] := 0.27214491;
      R_o[6,6] := -0.01843679;
      R_o[6,7] := 0.23837006;
      R_o[7,0] := 0.42624715;
      R_o[7,1] := 0.84213698;
      R_o[7,2] := 1.39297855;
      R_o[7,3] := 0.25695744;
      R_o[7,4] := -0.87713885;
      R_o[7,5] := -0.13476479;
      R_o[7,6] := -0.05455340;
      R_o[7,7] := 0.17162661;
      B_i[0] := 0.87045062;
      B_i[1] := 0.38770351;
      B_i[2] := -0.11886705;
      B_i[3] := -0.35644138;
      B_i[4] := -0.07135087;
      B_i[5] := 1.00623786;
      B_i[6] := 0.26473454;
      B_i[7] := 1.23754025;
      B_f[0] := 1.99891639;
      B_f[1] := 2.66124272;
      B_f[2] := 1.60180199;
      B_f[3] := 3.88835764;
      B_f[4] := 1.62835073;
      B_f[5] := 0.97422898;
      B_f[6] := 2.22533846;
      B_f[7] := 1.28588867;
      B_g[0] := 0.27844557;
      B_g[1] := 0.63931465;
      B_g[2] := 1.02911937;
      B_g[3] := -0.69296604;
      B_g[4] := -1.26938105;
      B_g[5] := 0.09129135;
      B_g[6] := -0.87523937;
      B_g[7] := -0.22564322;
      B_o[0] := 3.00663900;
      B_o[1] := 2.94506073;
      B_o[2] := 2.22459459;
      B_o[3] := 3.24792528;
      B_o[4] := 3.54929399;
      B_o[5] := 3.08820629;
      B_o[6] := 2.67632246;
      B_o[7] := 3.11170125;
      FC_W[0,0] := -1.37318242;
      FC_W[0,1] := -0.52894771;
      FC_W[0,2] := 0.82508540;
      FC_W[0,3] := -1.99275565;
      FC_W[0,4] := 1.18965185;
      FC_W[0,5] := 2.38302135;
      FC_W[0,6] := 0.24659581;
      FC_W[0,7] := 0.36538163;
      FC_W[1,0] := 0.27071670;
      FC_W[1,1] := 0.41951901;
      FC_W[1,2] := 1.60569334;
      FC_W[1,3] := 1.23515272;
      FC_W[1,4] := -2.97889638;
      FC_W[1,5] := -1.94566178;
      FC_W[1,6] := 0.43387899;
      FC_W[1,7] := 0.16437700;
      FC_W[2,0] := -1.35792935;
      FC_W[2,1] := -0.49226213;
      FC_W[2,2] := 0.80376226;
      FC_W[2,3] := -1.97948229;
      FC_W[2,4] := 1.19592011;
      FC_W[2,5] := 2.36552095;
      FC_W[2,6] := 0.23025335;
      FC_W[2,7] := 0.34811801;
      FC_W[3,0] := 0.68208855;
      FC_W[3,1] := 0.12471101;
      FC_W[3,2] := 0.07761292;
      FC_W[3,3] := -2.11483049;
      FC_W[3,4] := 1.25893140;
      FC_W[3,5] := 0.99728709;
      FC_W[3,6] := -1.82845187;
      FC_W[3,7] := -0.19247104;
      FC_W[4,0] := -1.44672430;
      FC_W[4,1] := -0.50926137;
      FC_W[4,2] := -2.30950522;
      FC_W[4,3] := -1.96016002;
      FC_W[4,4] := -0.92503679;
      FC_W[4,5] := -1.26670945;
      FC_W[4,6] := -0.08506308;
      FC_W[4,7] := 0.52047390;
      FC_W[5,0] := 0.44260150;
      FC_W[5,1] := 0.37026632;
      FC_W[5,2] := 1.35409307;
      FC_W[5,3] := 0.15279016;
      FC_W[5,4] := 0.37467703;
      FC_W[5,5] := -0.87928665;
      FC_W[5,6] := 1.43426895;
      FC_W[5,7] := 0.70363981;
      FC_W[6,0] := 1.77307248;
      FC_W[6,1] := -0.50528181;
      FC_W[6,2] := 0.85060036;
      FC_W[6,3] := -1.50316060;
      FC_W[6,4] := 1.24707830;
      FC_W[6,5] := -0.39548868;
      FC_W[6,6] := 1.74957681;
      FC_W[6,7] := -0.27180871;
      FC_W[7,0] := 0.66992402;
      FC_W[7,1] := 0.10731039;
      FC_W[7,2] := 0.07762623;
      FC_W[7,3] := -2.13342810;
      FC_W[7,4] := 1.26615632;
      FC_W[7,5] := 1.01499653;
      FC_W[7,6] := -1.81981516;
      FC_W[7,7] := -0.17927456;
      FC_W[8,0] := 0.66936851;
      FC_W[8,1] := 0.14543790;
      FC_W[8,2] := 0.03346241;
      FC_W[8,3] := -2.01580858;
      FC_W[8,4] := 1.34549654;
      FC_W[8,5] := 0.98734695;
      FC_W[8,6] := -1.81929374;
      FC_W[8,7] := -0.16405965;
      FC_W[9,0] := 0.66745198;
      FC_W[9,1] := 0.12200294;
      FC_W[9,2] := 0.08669009;
      FC_W[9,3] := -2.12185860;
      FC_W[9,4] := 1.27060866;
      FC_W[9,5] := 1.02163804;
      FC_W[9,6] := -1.83411348;
      FC_W[9,7] := -0.17880493;
      FC_W[10,0] := -0.43640897;
      FC_W[10,1] := 0.68268049;
      FC_W[10,2] := 0.14224736;
      FC_W[10,3] := -0.68086797;
      FC_W[10,4] := 0.35580847;
      FC_W[10,5] := 0.92224455;
      FC_W[10,6] := -2.43797994;
      FC_W[10,7] := 0.26598689;
      FC_W[11,0] := 0.35488737;
      FC_W[11,1] := 1.68916869;
      FC_W[11,2] := -1.16505313;
      FC_W[11,3] := -1.03148413;
      FC_W[11,4] := -0.62006569;
      FC_W[11,5] := 0.32353073;
      FC_W[11,6] := 0.20904805;
      FC_W[11,7] := -1.50123751;
      FC_W[12,0] := 0.75137240;
      FC_W[12,1] := 1.51158011;
      FC_W[12,2] := -0.97034442;
      FC_W[12,3] := -1.03762329;
      FC_W[12,4] := -0.62972116;
      FC_W[12,5] := 0.15404159;
      FC_W[12,6] := -0.13045871;
      FC_W[12,7] := -1.14926791;
      FC_W[13,0] := -1.24091721;
      FC_W[13,1] := 0.72264183;
      FC_W[13,2] := 4.21143913;
      FC_W[13,3] := -0.64818949;
      FC_W[13,4] := -2.22882915;
      FC_W[13,5] := 0.28011763;
      FC_W[13,6] := 0.08918135;
      FC_W[13,7] := 1.46233487;
      FC_W[14,0] := -1.83078206;
      FC_W[14,1] := -1.94626880;
      FC_W[14,2] := 2.02099109;
      FC_W[14,3] := -0.88200986;
      FC_W[14,4] := 1.19228423;
      FC_W[14,5] := -2.04054785;
      FC_W[14,6] := -1.13131750;
      FC_W[14,7] := -3.02692223;
      FC_W[15,0] := -0.17234646;
      FC_W[15,1] := 1.68070006;
      FC_W[15,2] := -0.98812079;
      FC_W[15,3] := -1.02355719;
      FC_W[15,4] := -0.51346064;
      FC_W[15,5] := 0.30412915;
      FC_W[15,6] := 0.49580911;
      FC_W[15,7] := -2.00975895;
      FC_W[16,0] := 0.14178839;
      FC_W[16,1] := -2.42272043;
      FC_W[16,2] := 1.82622004;
      FC_W[16,3] := -0.81107336;
      FC_W[16,4] := 1.03681660;
      FC_W[16,5] := -1.79800606;
      FC_W[16,6] := -2.25264025;
      FC_W[16,7] := -0.61567187;
      FC_W[17,0] := 3.12230635;
      FC_W[17,1] := -1.14041483;
      FC_W[17,2] := 0.45076677;
      FC_W[17,3] := 0.17650086;
      FC_W[17,4] := -0.00877836;
      FC_W[17,5] := -0.71208066;
      FC_W[17,6] := -2.28671813;
      FC_W[17,7] := 3.42369246;
      FC_W[18,0] := 0.76313448;
      FC_W[18,1] := -1.93009770;
      FC_W[18,2] := -4.29185629;
      FC_W[18,3] := -1.50427651;
      FC_W[18,4] := -0.13721293;
      FC_W[18,5] := 0.55832797;
      FC_W[18,6] := 0.58232069;
      FC_W[18,7] := -1.97768271;
      FC_W[19,0] := 0.58457559;
      FC_W[19,1] := 1.94365251;
      FC_W[19,2] := -0.06313096;
      FC_W[19,3] := -0.65289688;
      FC_W[19,4] := -0.60565686;
      FC_W[19,5] := 0.01970079;
      FC_W[19,6] := -0.15449062;
      FC_W[19,7] := -0.71010417;
      FC_W[20,0] := -1.53441155;
      FC_W[20,1] := 0.26765692;
      FC_W[20,2] := -0.60537034;
      FC_W[20,3] := 0.46610016;
      FC_W[20,4] := -1.96675193;
      FC_W[20,5] := 0.30353904;
      FC_W[20,6] := -1.85867703;
      FC_W[20,7] := 0.08975823;
      FC_W[21,0] := 2.47608876;
      FC_W[21,1] := -1.64168596;
      FC_W[21,2] := -0.25707519;
      FC_W[21,3] := -1.46445429;
      FC_W[21,4] := -0.22880352;
      FC_W[21,5] := 1.31707644;
      FC_W[21,6] := 0.93424761;
      FC_W[21,7] := -2.32273722;
      FC_W[22,0] := 0.52312243;
      FC_W[22,1] := -0.79484791;
      FC_W[22,2] := 2.66410828;
      FC_W[22,3] := -3.21130037;
      FC_W[22,4] := -4.10494614;
      FC_W[22,5] := -0.08404513;
      FC_W[22,6] := -0.47616670;
      FC_W[22,7] := -0.67225242;
      FC_W[23,0] := -1.20075583;
      FC_W[23,1] := 1.00352490;
      FC_W[23,2] := 4.44261217;
      FC_W[23,3] := -1.13683903;
      FC_W[23,4] := -1.55746245;
      FC_W[23,5] := 0.62567723;
      FC_W[23,6] := -0.98258156;
      FC_W[23,7] := 1.32669258;
      FC_W[24,0] := 0.58476400;
      FC_W[24,1] := -0.88437301;
      FC_W[24,2] := 2.53204155;
      FC_W[24,3] := -3.27082038;
      FC_W[24,4] := -4.12127066;
      FC_W[24,5] := -0.07652019;
      FC_W[24,6] := -0.42923889;
      FC_W[24,7] := -0.77052402;
      FC_W[25,0] := 0.58642721;
      FC_W[25,1] := -0.88521427;
      FC_W[25,2] := 2.53265524;
      FC_W[25,3] := -3.27612162;
      FC_W[25,4] := -4.12974119;
      FC_W[25,5] := -0.07558586;
      FC_W[25,6] := -0.42920873;
      FC_W[25,7] := -0.77160281;
      FC_W[26,0] := -1.19534051;
      FC_W[26,1] := 0.86386824;
      FC_W[26,2] := 3.25430202;
      FC_W[26,3] := -1.30819666;
      FC_W[26,4] := -2.58638358;
      FC_W[26,5] := -1.03585303;
      FC_W[26,6] := -0.78927201;
      FC_W[26,7] := 1.44714129;
      FC_W[27,0] := 2.27338052;
      FC_W[27,1] := -1.59377396;
      FC_W[27,2] := -0.89853072;
      FC_W[27,3] := -1.03837013;
      FC_W[27,4] := 0.30014247;
      FC_W[27,5] := 1.39629662;
      FC_W[27,6] := 0.90782219;
      FC_W[27,7] := -2.27797079;
      FC_W[28,0] := -0.92284089;
      FC_W[28,1] := 0.07467480;
      FC_W[28,2] := -0.87209713;
      FC_W[28,3] := -2.03417110;
      FC_W[28,4] := 0.61149502;
      FC_W[28,5] := -1.26839030;
      FC_W[28,6] := 1.43396020;
      FC_W[28,7] := 0.94821721;
      FC_W[29,0] := -0.58881819;
      FC_W[29,1] := 0.79866910;
      FC_W[29,2] := -2.62302852;
      FC_W[29,3] := 3.12394333;
      FC_W[29,4] := 3.99654388;
      FC_W[29,5] := 0.08908840;
      FC_W[29,6] := 0.47106421;
      FC_W[29,7] := 0.68441206;
      FC_W[30,0] := 0.51938868;
      FC_W[30,1] := -0.79148084;
      FC_W[30,2] := 2.66624427;
      FC_W[30,3] := -3.20863032;
      FC_W[30,4] := -4.10495043;
      FC_W[30,5] := -0.08509474;
      FC_W[30,6] := -0.47728243;
      FC_W[30,7] := -0.66817790;
      FC_W[31,0] := 0.49553028;
      FC_W[31,1] := -0.75901192;
      FC_W[31,2] := 2.68577194;
      FC_W[31,3] := -3.16863751;
      FC_W[31,4] := -4.06989050;
      FC_W[31,5] := -0.10302582;
      FC_W[31,6] := -0.47943082;
      FC_W[31,7] := -0.63844413;
      FC_W[32,0] := 0.61318892;
      FC_W[32,1] := -0.88193792;
      FC_W[32,2] := 2.58489490;
      FC_W[32,3] := -3.27777791;
      FC_W[32,4] := -4.12373161;
      FC_W[32,5] := -0.08388495;
      FC_W[32,6] := -0.41740480;
      FC_W[32,7] := -0.76095468;
      FC_W[33,0] := 0.61156529;
      FC_W[33,1] := -0.83659351;
      FC_W[33,2] := 2.64606047;
      FC_W[33,3] := -3.22972894;
      FC_W[33,4] := -4.07023621;
      FC_W[33,5] := -0.12561664;
      FC_W[33,6] := -0.41470754;
      FC_W[33,7] := -0.70742649;
      FC_W[34,0] := 0.56957924;
      FC_W[34,1] := -0.81484163;
      FC_W[34,2] := 2.66175270;
      FC_W[34,3] := -3.22360635;
      FC_W[34,4] := -4.08081150;
      FC_W[34,5] := -0.11388451;
      FC_W[34,6] := -0.44544184;
      FC_W[34,7] := -0.67890739;
      FC_W[35,0] := 0.62116420;
      FC_W[35,1] := -0.91804183;
      FC_W[35,2] := 2.55082273;
      FC_W[35,3] := -3.30127358;
      FC_W[35,4] := -4.12339067;
      FC_W[35,5] := -0.04686525;
      FC_W[35,6] := -0.41361472;
      FC_W[35,7] := -0.80192775;
      FC_W[36,0] := 0.96057558;
      FC_W[36,1] := -1.52714062;
      FC_W[36,2] := -0.09157373;
      FC_W[36,3] := -2.29993343;
      FC_W[36,4] := -2.74687934;
      FC_W[36,5] := 0.89486367;
      FC_W[36,6] := -0.21753848;
      FC_W[36,7] := -1.98280287;
      FC_W[37,0] := 0.63659966;
      FC_W[37,1] := -0.92864555;
      FC_W[37,2] := 2.55096030;
      FC_W[37,3] := -3.30504990;
      FC_W[37,4] := -4.11750746;
      FC_W[37,5] := -0.03328575;
      FC_W[37,6] := -0.40167740;
      FC_W[37,7] := -0.81976414;
      FC_W[38,0] := -1.57151544;
      FC_W[38,1] := -2.32424641;
      FC_W[38,2] := 2.13469505;
      FC_W[38,3] := -1.01246119;
      FC_W[38,4] := 1.27655017;
      FC_W[38,5] := -2.01633477;
      FC_W[38,6] := -1.49836993;
      FC_W[38,7] := -2.66122508;
      FC_W[39,0] := -1.85308564;
      FC_W[39,1] := -2.34909940;
      FC_W[39,2] := 2.25910854;
      FC_W[39,3] := -1.06350100;
      FC_W[39,4] := 1.33850765;
      FC_W[39,5] := -2.17299938;
      FC_W[39,6] := -1.42110384;
      FC_W[39,7] := -3.07338285;
      FC_B[0] := -0.03680599;
      FC_B[1] := -0.99531233;
      FC_B[2] := -0.03512276;
      FC_B[3] := -0.51894927;
      FC_B[4] := -0.34805626;
      FC_B[5] := -0.10473614;
      FC_B[6] := 0.16657342;
      FC_B[7] := -0.51048559;
      FC_B[8] := -0.46436945;
      FC_B[9] := -0.51502335;
      FC_B[10] := -0.66331333;
      FC_B[11] := -0.91201615;
      FC_B[12] := -0.94463032;
      FC_B[13] := -1.87086606;
      FC_B[14] := 0.51885176;
      FC_B[15] := -0.82386893;
      FC_B[16] := 0.42529055;
      FC_B[17] := -0.09486814;
      FC_B[18] := 1.10968602;
      FC_B[19] := -1.16007948;
      FC_B[20] := -0.65581632;
      FC_B[21] := 0.40555862;
      FC_B[22] := -2.37383127;
      FC_B[23] := -2.08129168;
      FC_B[24] := -2.33415413;
      FC_B[25] := -2.33819509;
      FC_B[26] := -2.22797513;
      FC_B[27] := 0.78016996;
      FC_B[28] := -0.22360271;
      FC_B[29] := 2.31837344;
      FC_B[30] := -2.37427068;
      FC_B[31] := -2.37652969;
      FC_B[32] := -2.34959030;
      FC_B[33] := -2.34812522;
      FC_B[34] := -2.36254501;
      FC_B[35] := -2.33670855;
      FC_B[36] := -0.85175836;
      FC_B[37] := -2.33044815;
      FC_B[38] := 0.57427269;
      FC_B[39] := 0.59669638;

END_DATA_BLOCK
